Fanuc KAREL source: kb00202.KL

-- PROVISIONAL review KL for V770-1; original PC SHA256 7e14280f9021a7437fc2b8b7f5d4fe01d7c69d6d1de910350c3ab9f3eb8ed3a3
-- Incomplete behavior may be omitted. Consult companion uncertainty JSON. Do not deploy.
PROGRAM KB00202
%NOLOCKGROUP
BEGIN
  -- UNRESOLVED_PC offsets 5-14; opcodes 3F,75
  -- UNRESOLVED_PC offsets 19-28; opcodes 3F,75
  -- UNRESOLVED_PC offsets 33-40; opcodes 9D,23
  -- UNRESOLVED_PC offsets 45-77; opcodes 27,22,22,2A,22,2A,22,31
  -- UNRESOLVED_PC offsets 82-86; opcodes 7F
END KB00202
